// TIA Portal V21 export
DATA_BLOCK "AxisAS_SimIO"   // DB900
{ S7_Optimized_Access := 'FALSE' }
VERSION : 0.1
// Scambio PLC <-> simulatore encoder AxisAS_Sim_v4.py (snap7). Accesso STANDARD: offset fissi, non modificare l'ordine.
// stored: AutoNumber false
   VAR
      xCmdForw : Bool := false;   // PLC -> SIM 0.0 Marcia avanti
      xCmdBack : Bool := false;   // PLC -> SIM 0.1 Marcia indietro
      xCmdBrake : Bool := false;   // PLC -> SIM 0.2 Sblocco freno
      fSpeedRef : Real := 0.0;   // PLC -> SIM 2 Riferimento velocità (mm/s, modulo)
      fEncoder : Real := 0.0;   // SIM -> PLC 6 Posizione encoder simulata (mm)
      xDriveReady : Bool := false;   // SIM -> PLC 10.0 Inverter pronto / magnetizzato
      xLevelSensor : Bool := false;   // SIM -> PLC 10.1 Sensore livello virtuale
      iHeartbeat : Int := 0;   // SIM -> PLC 12 Contatore vita del simulatore
   END_VAR
BEGIN
END_DATA_BLOCK
